(* IEC 61131-3 sources: SortJet_MasterSPS_Aufbau.fbsproj/12_Visu_Uebersicht, 12 files *)

(* ---- VISU_HAND.gvl ---- *)
(* METADATA
{
	"v3Meta": {
		"objectGuid": "6f32179b-dff3-42c9-9870-23893e477a6b"
	}
}
*)
{attribute 'qualified_only'}
NAMESPACE VISU_HAND
VAR_GLOBAL
  st201  : VisuHand_Station_ST;
  st202  : VisuHand_Station_ST;
  st203  : VisuHand_Station_ST;
  st204  : VisuHand_Station_ST;
  st205  : VisuHand_Station_ST;
  st206  : VisuHand_Station_ST;
  st207  : VisuHand_Station_ST;
  st208  : VisuHand_Station_ST;
  st101  : VisuHand_Station_ST;
  st102  : VisuHand_Station_ST;
  st151  : VisuHand_Station_ST;
  st152  : VisuHand_Station_ST;
  astFW  : ARRAY[301..305] OF VisuHand_Station_ST;

  bAnlageResetTaster : BOOL;          // Visu-Taster Anlagen-Reset (einfacher Druck)
  bAnlageResetAktiv  : BOOL;          // Reset laeuft (min. 1 s angezeigt, solange eine Station noch bReset hat)
  sAnlageReset       : STRING(40) := 'ANLAGE RESET';
  dwAnlageResetFarbe : DWORD := 16#FFD64545;
  sLblReset          : STRING(20) := 'Reset';

  // Beschriftungen der Visu "Handbetrieb" (benannt, damit Visu und GVL nicht unbemerkt auseinanderlaufen)
  sL_Riemen                                : STRING(120) := 'Riemen';
  sL_Riemen_X                              : STRING(120) := 'Riemen X';
  sL_Riemen_Y                              : STRING(120) := 'Riemen Y';
  sL_Zur_Zurueck                           : STRING(120) := '<< Zurück';
  sL_Vor_Vor                               : STRING(120) := 'Vor >>';
  sL_Anschlag                              : STRING(120) := 'Anschlag';
  sL_Ab                                    : STRING(120) := 'Ab';
  sL_Auf                                   : STRING(120) := 'Auf';
  sL_Hubrahmen                             : STRING(120) := 'Hubrahmen';
  sL_Senken                                : STRING(120) := 'Senken';
  sL_Heben                                 : STRING(120) := 'Heben';
  sL_Messachse                             : STRING(120) := 'Messachse';
  sL_Minus_Ab                              : STRING(120) := '- Ab';
  sL_Plus_Auf                              : STRING(120) := '+ Auf';
  sL_Referenz                              : STRING(120) := 'Referenz';
  sL_Geblaese                              : STRING(120) := 'Gebläse';
  sL_Ein_Aus                               : STRING(120) := 'Ein / Aus';
  sL_Drosselkl                             : STRING(120) := 'Drosselkl.';
  sL_Auf_Zu                                : STRING(120) := 'Auf / Zu';
  sL_Kippen                                : STRING(120) := 'Kippen';
  sL_Waagerecht                            : STRING(120) := 'Waagerecht';
  sL_Senkrecht                             : STRING(120) := 'Senkrecht';
  sL_Querfahrt                             : STRING(120) := 'Querfahrt';
  sL_Minus_Minus                           : STRING(120) := '- Minus';
  sL_Plus_Plus                             : STRING(120) := '+ Plus';
  sL_84Grad                                : STRING(120) := '84°';
  sL_90Grad                                : STRING(120) := '90°';
  sL_Schmierung                            : STRING(120) := 'Schmierung';
  sL_Starten                               : STRING(120) := 'Starten';
  sL_Riemen_Hub                            : STRING(120) := 'Riemen Hub';
  sL_Anheben                               : STRING(120) := 'Anheben';
  sL_Abfr_Einl                             : STRING(120) := 'Abfr. Einl.';
  sL_Luft_ein                              : STRING(120) := 'Luft ein';
  sL_Abfr_Ausl                             : STRING(120) := 'Abfr. Ausl.';
  sL_Rolltor                               : STRING(120) := 'Rolltor';
  sL_Runter                                : STRING(120) := 'Runter';
  sL_Hoch                                  : STRING(120) := 'Hoch';
  sL_Linearein                             : STRING(120) := 'Linearein.';
  sL_Zurueck                               : STRING(120) := 'Zurück';
  sL_Vor                                   : STRING(120) := 'Vor';
  sL_Shuttle                               : STRING(120) := 'Shuttle';
  sL_Greifer                               : STRING(120) := 'Greifer';
  sL_Oeffnen                               : STRING(120) := 'Öffnen';
  sL_Schliessen                            : STRING(120) := 'Schließen';
  sL_Entriegel                             : STRING(120) := 'Entriegel.';
  sL_Gegenhalter                           : STRING(120) := 'Gegenhalter';
  sL_Lichtschr                             : STRING(120) := 'Lichtschr.';
  sL_Quittieren                            : STRING(120) := 'Quittieren';
  sL_Oeffnung                              : STRING(120) := 'Öffnung';
  sL_16mm                                  : STRING(120) := '16 mm';
  sL_23mm                                  : STRING(120) := '23 mm';
  sL_29mm                                  : STRING(120) := '29 mm';
  sL_Greiferachse                          : STRING(120) := 'Gr.-Achse';
  sL_Zange                                 : STRING(120) := 'Zange';
  sL_Rueckhalter                           : STRING(120) := 'Rückhalter';
  sL_Drehen                                : STRING(120) := 'Drehen';
  sL_0Grad                                 : STRING(120) := '0°';
  sL_180Grad                               : STRING(120) := '180°';
  sL_270Grad                               : STRING(120) := '270°';
  sL_Arretierung                           : STRING(120) := 'Arretierung';
  sL_Einfahren                             : STRING(120) := 'Einfahren';
  sL_Ausfahren                             : STRING(120) := 'Ausfahren';
  sL_Abschrankung                          : STRING(120) := 'Abschrank.';
  sL_HANDBETRIEB                           : STRING(120) := 'HANDBETRIEB';
  sL_Legende                               : STRING(120) := 'Taster (weiß) = Tippbetrieb solange gedrückt   |   Schalter (blau hinterlegt wenn EIN) = Ein/Aus   |   Gesperrt = grau';
  sL_Titel                                 : STRING(120) := 'SortJet  -  Handbetrieb 201 - 208';
  sL_Titel2                                : STRING(120) := 'SortJet  -  Handbetrieb Speicher';
END_VAR
END_NAMESPACE

(* ---- VISU_UEBERSICHT.gvl ---- *)
(* METADATA
{
	"v3Meta": {
		"objectGuid": "76464f8f-3613-4465-9c50-3e0a0f70c8ba"
	}
}
*)
{attribute 'qualified_only'}
NAMESPACE VISU_UEBERSICHT
VAR_GLOBAL
  // Kopfzeile / Anlagenstatus
  sTitel            : STRING(80) := 'SortJet -  Anlagenübersicht';
  sUntertitel       : STRING(120) := 'Anlegetisch 201/205 > Eckübergabe 204 > Drehstation 207 > Shuttle 101 > Speicher > Shuttle 102 > Fächerwagen';
  stAutomatik       : VisuUeb_Lampe_ST;
  stSK1             : VisuUeb_Lampe_ST;
  stSK2             : VisuUeb_Lampe_ST;
  stSK3             : VisuUeb_Lampe_ST;
  stSK4             : VisuUeb_Lampe_ST;
  astTuer               : ARRAY[1..cMAX_TUEREN] OF VisuUeb_Lampe_ST;      // je Tuer eine Anzeige
  abTuerVorhanden       : ARRAY[1..cMAX_TUEREN] OF BOOL;
  astDurchgang          : ARRAY[1..cMAX_DURCHGAENGE] OF VisuUeb_Lampe_ST;
  abDurchgangVorhanden  : ARRAY[1..cMAX_DURCHGAENGE] OF BOOL;
  sLblTueren            : STRING(20) := 'TÜREN';
  sLblDurchgaenge       : STRING(20) := 'DURCHGÄNGE';
  stDruckluft       : VisuUeb_Lampe_ST;
  stSchaltschrank   : VisuUeb_Lampe_ST;
  stEtherCAT        : VisuUeb_Lampe_ST;
  stInit            : VisuUeb_Lampe_ST;
  stMMI             : VisuUeb_Lampe_ST;
  stBetriebsstop    : VisuUeb_Lampe_ST;
  stInbetriebnahme  : VisuUeb_Lampe_ST;
  sStoerungen       : STRING(80);
  dwStoerungenFarbe : DWORD := 16#FF2EAD5B;

  // Stationen
  st501             : VisuUeb_Station_ST;
  st201             : VisuUeb_Station_ST;
  st202             : VisuUeb_Station_ST;
  st203             : VisuUeb_Station_ST;
  st204             : VisuUeb_Station_ST;
  st205             : VisuUeb_Station_ST;
  st206             : VisuUeb_Station_ST;
  st207             : VisuUeb_Station_ST;
  st208             : VisuUeb_Station_ST;
  st101             : VisuUeb_Station_ST;
  st102             : VisuUeb_Station_ST;
  st151             : VisuUeb_Station_ST;
  st152             : VisuUeb_Station_ST;
  st301             : VisuUeb_Station_ST;
  st302             : VisuUeb_Station_ST;
  st303             : VisuUeb_Station_ST;
  st304             : VisuUeb_Station_ST;
  st305             : VisuUeb_Station_ST;

  // Achsen (Querfahrt)
  stAchse101        : VisuUeb_Achse_ST;
  stAchse102        : VisuUeb_Achse_ST;
  stAchse151        : VisuUeb_Achse_ST;
  stAchse152        : VisuUeb_Achse_ST;

  // feste Beschriftungen (Visu nutzt ausschließlich Textvariablen)
  sLblSensoren      : STRING(40) := 'E       EV      AV       A';
  sLblSpeicher      : STRING(40) := 'S O R T I E R S P E I C H E R';
  sLblShuttle101    : STRING(40) := 'SHUTTLE 101';
  sLblTS151         : STRING(40) := 'TRANSFERSHUTTLE 151';
  sLblReset         : STRING(40) := 'Skalierung neu lernen';
  sLblLegende       : STRING(120) := 'Grün = Automatik    Orange = Hand    Blau = Reset / Referenz    Rot = Störung    Grau = deaktiviert';
  sLblNotHaltOK     : STRING(40) := 'NOT-HALT OK';
  sLblNotHaltAus    : STRING(40) := 'NOT-HALT AUSGELÖST';
  sLblStatus        : STRING(40) := 'ANLAGENSTATUS';
  sLblQuerfahrt     : STRING(40) := 'QUERFAHRT';
  sLblIst           : STRING(20) := 'Ist';
  sLblZiel          : STRING(20) := 'Ziel';
  sLblSpeed         : STRING(20) := 'v';
  sLblE             : STRING(4)  := 'E';
  sLblEV            : STRING(4)  := 'EV';
  sLblAV            : STRING(4)  := 'AV';
  sLblA             : STRING(4)  := 'A';
  sLblAS            : STRING(4)  := 'AS';
  sLblQuer101       : STRING(60) := 'QUERFAHRT SHUTTLE 101';
  sLblQuer102       : STRING(60) := 'QUERFAHRT SHUTTLE 102';
  sLblWagen101      : STRING(20) := '101';
  sLblWagen102      : STRING(20) := '102';
  sLblZielMarke     : STRING(10) := 'ZIEL';

  // Bedienung
  bSkalierungNeuLernen : BOOL;
END_VAR

VAR_GLOBAL RETAIN
  // Selbstlernende Skalierung der Fahrbahnen (min/max beobachtete Position)
  bSkalierung101Init : BOOL;
  rMin101            : REAL;
  rMax101            : REAL;
  bSkalierung102Init : BOOL;
  rMin102            : REAL;
  rMax102            : REAL;
  bSkalierung151Init : BOOL;
  rMin151            : REAL;
  rMax151            : REAL;
  bSkalierung152Init : BOOL;
  rMin152            : REAL;
  rMax152            : REAL;
END_VAR

VAR_GLOBAL CONSTANT
  cMAX_TUEREN          : WORD := 8;     // Anzahl Tueranzeigen in der Visu
  cMAX_DURCHGAENGE     : WORD := 3;     // Anzahl Durchganganzeigen in der Visu
  cBAHN_LAENGE_PX      : INT  := 266;   // nutzbare Laenge der senkrechten Fahrbahn (muss zur Visu passen)
  cWAGEN_LAENGE_PX     : INT  := 34;    // Hoehe Fahrwagen (muss zur Visu passen)
  cMIN_SPANNE_MM       : REAL := 500;   // minimale Skalierungsspanne

  cFARBE_GRUEN         : DWORD := 16#FF2EAD5B;
  cFARBE_ROT           : DWORD := 16#FFD64545;
  cFARBE_ORANGE        : DWORD := 16#FFF0A202;
  cFARBE_BLAU          : DWORD := 16#FF2F80ED;
  cFARBE_GRAU          : DWORD := 16#FF9AA5B1;
  cFARBE_GRAU_HELL     : DWORD := 16#FFE4E7EB;
  cFARBE_RAHMEN        : DWORD := 16#FFCBD2D9;
  cFARBE_TEXT          : DWORD := 16#FF52606D;
  cFARBE_SENSOR_AN     : DWORD := 16#FFFFC531;
END_VAR
END_NAMESPACE

(* ---- VisuHand_Set.fn.st ---- *)
(* METADATA
{
	"v3Meta": {
		"objectGuid": "443bc09b-b8af-4511-9c3a-ed00ec4cc080"
	}
}
*)
FUNCTION VisuHand_Set : BOOL
VAR_IN_OUT
  stH     : VisuHand_Station_ST;
END_VAR
VAR_INPUT
  wZeile  : WORD;
  sText   : STRING(30);
  dwFarbe : DWORD;
END_VAR
IF wZeile >= 1 AND wZeile <= 10 THEN // Grenzen wie VisuHand_Station_ST.asStatus
  stH.asStatus[wZeile]  := sText;
  stH.adwStatus[wZeile] := dwFarbe;
END_IF
VisuHand_Set := TRUE;
END_FUNCTION

(* ---- VisuHand_Sperre.fn.st ---- *)
(* METADATA
{
	"v3Meta": {
		"objectGuid": "d31da620-9df0-4563-ab06-3d7039f98cd3"
	}
}
*)
FUNCTION VisuHand_Sperre : BOOL
VAR_IN_OUT
  stBP : StationBasisParameter_ST;
  stH  : VisuHand_Station_ST;
END_VAR
VAR_INPUT
  bFaecherwagen : BOOL; // FW-Handfunktionen sind im FB nicht an die Betriebsart gebunden -> hier zusaetzlich bei Automatik sperren
END_VAR
VAR
  bDeaktiviert : BOOL;
END_VAR
IF __ISVALIDREF(stBP.stMKs) THEN
  bDeaktiviert := stBP.stMKs.bDeaktivieren;
END_IF

IF bDeaktiviert THEN
  stH.bGesperrt := TRUE;  stH.sSperrgrund := 'Gesperrt: Station deaktiviert';
ELSIF stBP.bAutomatik THEN
  stH.bGesperrt := TRUE;  stH.sSperrgrund := 'Gesperrt: Automatik aktiv';
ELSIF stBP.bReset THEN
  stH.bGesperrt := TRUE;  stH.sSperrgrund := 'Gesperrt: Reset läuft';
ELSIF stBP.bReferenz THEN
  stH.bGesperrt := TRUE;  stH.sSperrgrund := 'Gesperrt: Referenzfahrt läuft';
ELSIF stBP.bCheck THEN
  stH.bGesperrt := TRUE;  stH.sSperrgrund := 'Gesperrt: Systemcheck läuft';
ELSIF bFaecherwagen AND (stBP.bEintransport[cWAND_1] OR stBP.bAustransport[cWAND_1]) THEN
  stH.bGesperrt := TRUE;  stH.sSperrgrund := 'Gesperrt: Ein-/Ausschleusen aktiv';
ELSE
  stH.bGesperrt := FALSE;
  stH.sSperrgrund := SEL(stBP.stFreigabe.bAlles, 'Hand frei - keine Sicherheitsfreigabe', 'Handbetrieb freigegeben');
END_IF

IF stH.bGesperrt THEN
  stH.dwSperrFarbe := VISU_UEBERSICHT.cFARBE_GRAU;
ELSIF NOT stBP.stFreigabe.bAlles THEN
  stH.dwSperrFarbe := VISU_UEBERSICHT.cFARBE_ORANGE;
ELSE
  stH.dwSperrFarbe := VISU_UEBERSICHT.cFARBE_GRUEN;
END_IF
VisuHand_Sperre := stH.bGesperrt;
END_FUNCTION

(* ---- VisuUeb_Achse.fn.st ---- *)
(* METADATA
{
	"v3Meta": {
		"objectGuid": "3979691c-e077-4914-8fb4-604417bd71fb"
	}
}
*)
FUNCTION VisuUeb_Achse : BOOL
VAR_IN_OUT
  stAchse   : VisuUeb_Achse_ST;
  bInit     : BOOL;  // Skalierung initialisiert (RETAIN)
  rMin      : REAL;  // gelerntes Minimum (RETAIN)
  rMax      : REAL;  // gelerntes Maximum (RETAIN)
END_VAR
VAR_INPUT
  rIst         : REAL;
  rZiel        : REAL;
  rSpeed       : REAL;
  bPositionierung : BOOL;
  bReferenziert   : BOOL;
  bFehler         : BOOL;
  bMinEnd         : BOOL;
  bMaxEnd         : BOOL;
  bNeuLernen      : BOOL;
  bBlink          : BOOL;
  rSkalaMin       : REAL;  // gemeinsamer Darstellungsbereich mehrerer Achsen (Max <= Min: eigener Bereich)
  rSkalaMax       : REAL;
END_VAR
VAR
  rSpanne : REAL;
  rFaktor : REAL;
  iWeg    : INT;
  rDarstMin : REAL;
END_VAR
// Skalierung lernen (nur mit gueltiger Referenz)
IF bNeuLernen THEN
  bInit := FALSE;
END_IF
IF bReferenziert THEN
  IF NOT bInit THEN
    rMin  := rIst;
    rMax  := rIst;
    bInit := TRUE;
  END_IF
  rMin := MIN(rMin, rIst);
  rMax := MAX(rMax, rIst);
  IF bPositionierung THEN
    rMin := MIN(rMin, rZiel);
    rMax := MAX(rMax, rZiel);
  END_IF
END_IF

IF rSkalaMax > rSkalaMin THEN
  rDarstMin := rSkalaMin;
  rSpanne   := MAX(rSkalaMax - rSkalaMin, VISU_UEBERSICHT.cMIN_SPANNE_MM);
ELSE
  rDarstMin := rMin;
  rSpanne   := MAX(rMax - rMin, VISU_UEBERSICHT.cMIN_SPANNE_MM);
END_IF
iWeg    := VISU_UEBERSICHT.cBAHN_LAENGE_PX - VISU_UEBERSICHT.cWAGEN_LAENGE_PX;

rFaktor := LIMIT(0.0, (rIst - rDarstMin) / rSpanne, 1.0);
stAchse.iPixel := REAL_TO_INT(rFaktor * INT_TO_REAL(iWeg));
rFaktor := LIMIT(0.0, (rZiel - rDarstMin) / rSpanne, 1.0);
stAchse.iZielPixel := REAL_TO_INT(rFaktor * INT_TO_REAL(iWeg));

stAchse.rIstPos         := rIst;
stAchse.rZielPos        := rZiel;
stAchse.rSpeed          := rSpeed;
stAchse.bPositionierung := bPositionierung;
stAchse.bReferenziert   := bReferenziert;
stAchse.sIstPos         := VisuUeb_MmText(sPrefix := 'Ist  ', rWert := rIst);
stAchse.sZielPos        := SEL(bPositionierung, 'Ziel  -', VisuUeb_MmText(sPrefix := 'Ziel  ', rWert := rZiel));
stAchse.sSpeed          := VisuUeb_MmText(sPrefix := 'v  ', rWert := rSpeed, sEinheit := ' mm/s');
stAchse.sBereich        := CONCAT(CONCAT(VisuUeb_MmText(sPrefix := 'Bereich ', rWert := rMin), ' ... '), VisuUeb_MmText(sPrefix := '', rWert := rMax));

IF bFehler THEN
  stAchse.dwKoerperFarbe := SEL(bBlink, 16#FF8C2F2F, VISU_UEBERSICHT.cFARBE_ROT);
ELSIF NOT bReferenziert THEN
  stAchse.dwKoerperFarbe := VISU_UEBERSICHT.cFARBE_ORANGE;
ELSIF bPositionierung THEN
  stAchse.dwKoerperFarbe := 16#FF1C64CC;
ELSE
  stAchse.dwKoerperFarbe := VISU_UEBERSICHT.cFARBE_BLAU;
END_IF
stAchse.dwMinEndFarbe := SEL(bMinEnd, VISU_UEBERSICHT.cFARBE_GRAU_HELL, VISU_UEBERSICHT.cFARBE_ROT);
stAchse.dwMaxEndFarbe := SEL(bMaxEnd, VISU_UEBERSICHT.cFARBE_GRAU_HELL, VISU_UEBERSICHT.cFARBE_ROT);
VisuUeb_Achse := bInit;
END_FUNCTION

(* ---- VisuUeb_Lampe.fn.st ---- *)
(* METADATA
{
	"v3Meta": {
		"objectGuid": "b7aa09e8-5cde-43cf-b09b-dc0ab15a15f2"
	}
}
*)
FUNCTION VisuUeb_Lampe : BOOL
VAR_IN_OUT
  stLampe   : VisuUeb_Lampe_ST;
END_VAR
VAR_INPUT
  sText     : STRING(40);
  bOK       : BOOL;   // TRUE = gruen
  bWarnung  : BOOL := FALSE; // bei NOT bOK: TRUE = orange, FALSE = rot
  bNeutral  : BOOL := FALSE; // TRUE = grau (inaktiv, keine Bewertung)
END_VAR
stLampe.sText := sText;
IF bNeutral THEN
  stLampe.dwFarbe := VISU_UEBERSICHT.cFARBE_GRAU;
ELSIF bOK THEN
  stLampe.dwFarbe := VISU_UEBERSICHT.cFARBE_GRUEN;
ELSIF bWarnung THEN
  stLampe.dwFarbe := VISU_UEBERSICHT.cFARBE_ORANGE;
ELSE
  stLampe.dwFarbe := VISU_UEBERSICHT.cFARBE_ROT;
END_IF
VisuUeb_Lampe := bOK;
END_FUNCTION

(* ---- VisuUeb_MmText.fn.st ---- *)
(* METADATA
{
	"v3Meta": {
		"objectGuid": "478effab-2bb6-4cba-a63b-7b7e6c506f75"
	}
}
*)
FUNCTION VisuUeb_MmText : STRING(40)
VAR_INPUT
  sPrefix : STRING(20);
  rWert   : REAL;
  sEinheit: STRING(10) := ' mm';
END_VAR
VisuUeb_MmText := CONCAT(CONCAT(sPrefix, DINT_TO_STRING(REAL_TO_DINT(rWert))), sEinheit);
END_FUNCTION

(* ---- VisuUeb_Sensor.fn.st ---- *)
(* METADATA
{
	"v3Meta": {
		"objectGuid": "2f1f2564-8eff-43f7-8c8f-4a939be6a082"
	}
}
*)
FUNCTION VisuUeb_Sensor : DWORD
VAR_INPUT
  bBelegt    : BOOL;
  bVorhanden : BOOL := TRUE;
END_VAR
IF NOT bVorhanden THEN
  VisuUeb_Sensor := 16#00FFFFFF; // transparent
ELSIF bBelegt THEN
  VisuUeb_Sensor := VISU_UEBERSICHT.cFARBE_SENSOR_AN;
ELSE
  VisuUeb_Sensor := VISU_UEBERSICHT.cFARBE_GRAU_HELL;
END_IF
END_FUNCTION

(* ---- VisuUeb_Station.fn.st ---- *)
(* METADATA
{
	"v3Meta": {
		"objectGuid": "2a69d02d-507f-4a31-bfce-f3b7167a1195"
	}
}
*)
FUNCTION VisuUeb_Station : BOOL
VAR_IN_OUT
  stBP    : StationBasisParameter_ST;
  stKarte : VisuUeb_Station_ST;
END_VAR
VAR_INPUT
  sTitel  : STRING(40);
  bBlink  : BOOL;
  bGlasZusatz : BOOL := FALSE; // zusaetzliche Glaserkennung (z.B. Sensoren)
  bReferenzRelevant : BOOL := TRUE; // FALSE: Station hat keine referenzierbaren Achsen (z.B. Faecherwagen)
END_VAR
VAR
  bDeaktiviert : BOOL;
END_VAR
stKarte.sTitel := sTitel;
IF __ISVALIDREF(stBP.stMKs) THEN
  bDeaktiviert := stBP.stMKs.bDeaktivieren;
END_IF
stKarte.bDeaktiviert := bDeaktiviert;

// Referenzstatus (BasisStationsParameter.bIstReferenziert)
stKarte.bReferenzAnzeigen := bReferenzRelevant AND NOT bDeaktiviert;
IF stBP.bIstReferenziert THEN
  stKarte.sReferenz := 'REFERENZIERT';      stKarte.dwReferenzFarbe := VISU_UEBERSICHT.cFARBE_GRUEN;
ELSIF stBP.bReferenz THEN
  stKarte.sReferenz := 'REFERENZIERT ...';  stKarte.dwReferenzFarbe := SEL(bBlink, VISU_UEBERSICHT.cFARBE_GRAU, VISU_UEBERSICHT.cFARBE_BLAU);
ELSE
  stKarte.sReferenz := 'NICHT REFERENZIERT'; stKarte.dwReferenzFarbe := VISU_UEBERSICHT.cFARBE_ORANGE;
END_IF

// Zustand
IF bDeaktiviert THEN
  stKarte.sZustand := 'DEAKTIVIERT';         stKarte.dwZustandFarbe := VISU_UEBERSICHT.cFARBE_GRAU;
ELSIF stBP.bFehler THEN
  stKarte.sZustand := 'STÖRUNG';             stKarte.dwZustandFarbe := VISU_UEBERSICHT.cFARBE_ROT;
ELSIF stBP.bReset THEN
  stKarte.sZustand := 'RESET';               stKarte.dwZustandFarbe := VISU_UEBERSICHT.cFARBE_BLAU;
ELSIF stBP.bReferenz THEN
  stKarte.sZustand := 'REFERENZFAHRT';       stKarte.dwZustandFarbe := VISU_UEBERSICHT.cFARBE_BLAU;
ELSIF stBP.bCheck THEN
  stKarte.sZustand := 'SYSTEMCHECK';         stKarte.dwZustandFarbe := VISU_UEBERSICHT.cFARBE_BLAU;
ELSIF stBP.bAutomatik THEN
  stKarte.sZustand := 'AUTOMATIK';           stKarte.dwZustandFarbe := VISU_UEBERSICHT.cFARBE_GRUEN;
ELSE
  stKarte.sZustand := 'HAND';                stKarte.dwZustandFarbe := VISU_UEBERSICHT.cFARBE_ORANGE;
END_IF

// Rahmen: Stoerung blinkt rot, aktiver Auftrag blau
IF stBP.bFehler AND NOT bDeaktiviert THEN
  stKarte.dwRahmenFarbe := SEL(bBlink, VISU_UEBERSICHT.cFARBE_RAHMEN, VISU_UEBERSICHT.cFARBE_ROT);
ELSIF stBP.bAuftragAktiv THEN
  stKarte.dwRahmenFarbe := VISU_UEBERSICHT.cFARBE_BLAU;
ELSE
  stKarte.dwRahmenFarbe := VISU_UEBERSICHT.cFARBE_RAHMEN;
END_IF

// Aktive Funktion
IF bDeaktiviert THEN
  stKarte.sFunktion := '-';
ELSIF stBP.bFehler THEN
  stKarte.sFunktion := CONCAT('Fehlernummer ', WORD_TO_STRING(stBP.wFehlerNummer));
ELSIF stBP.bAnlegen THEN                      stKarte.sFunktion := 'Anlegen';
ELSIF stBP.bAbnehmen THEN                     stKarte.sFunktion := 'Abnehmen';
ELSIF stBP.bEintransport[cWAND_1] THEN        stKarte.sFunktion := 'Eintransport';
ELSIF stBP.bAustransport[cWAND_1] THEN        stKarte.sFunktion := 'Austransport';
ELSIF stBP.bDurchtransport[cWAND_1] THEN      stKarte.sFunktion := 'Durchtransport';
ELSIF stBP.bVortransport[cWAND_1] THEN        stKarte.sFunktion := 'Vortransport';
ELSIF stBP.bTransportkopplung[cWAND_1] THEN   stKarte.sFunktion := 'Transportkopplung';
ELSIF stBP.bMesskopplung[cWAND_1] THEN        stKarte.sFunktion := 'Messkopplung';
ELSIF stBP.bGlaslaengenmessung THEN           stKarte.sFunktion := 'Glaslängenmessung';
ELSIF stBP.bGlashoehenmessung THEN            stKarte.sFunktion := 'Glashöhenmessung';
ELSIF stBP.bVorabpositionieren THEN           stKarte.sFunktion := 'Vorabpositionierung';
ELSIF stBP.bAuftragAktiv THEN                 stKarte.sFunktion := 'Auftrag aktiv';
ELSIF stBP.stFreigabe.bAlles THEN                     stKarte.sFunktion := 'Bereit';
ELSE                                          stKarte.sFunktion := 'Keine Freigabe';
END_IF

stKarte.bGlas := stBP.bStationBelegt[cWAND_1] OR bGlasZusatz;
VisuUeb_Station := stBP.bFehler AND NOT bDeaktiviert;
END_FUNCTION

(* ---- VisuHand_Reset_FB.fb.st ---- *)
(* METADATA
{
	"v3Meta": {
		"objectGuid": "8e79010e-8dea-435f-8304-0b4307ea198e"
	}
}
*)
FUNCTION_BLOCK VisuHand_Reset_FB
// Stations-Reset aus der Visu:
//   - setzt BasisStationsParameter.bReset (die Station fuehrt ihre eigene Reset-Aktion aus und setzt bReset selbst zurueck)
//   - nur ausserhalb der Automatik, nicht wenn die Station deaktiviert ist oder bereits ein Reset laeuft
VAR_IN_OUT
  stBP : StationBasisParameter_ST;
  stH  : VisuHand_Station_ST;
END_VAR
VAR
  rtlTaster    : R_TRIG;
  bDeaktiviert : BOOL;
END_VAR
bDeaktiviert := FALSE;
IF __ISVALIDREF(stBP.stMKs) THEN
  bDeaktiviert := stBP.stMKs.bDeaktivieren;
END_IF

stH.bResetGesperrt := bDeaktiviert OR stBP.bAutomatik OR stBP.bReset OR stBP.bReferenz OR stBP.bCheck;

rtlTaster(CLK := stH.bResetTaster);
IF rtlTaster.Q AND NOT stH.bResetGesperrt THEN
  stBP.bReset := TRUE;
END_IF
END_FUNCTION_BLOCK

(* ---- VisuHand_PRG.prg.st ---- *)
(* METADATA
{
	"v3Meta": {
		"objectGuid": "a4fab899-80a6-4d8b-aad2-f00973a33795"
	}
}
*)
PROGRAM VisuHand_PRG
VAR
  b    : BOOL;
  i    : WORD;
  dwG, dwO, dwR, dwGR, dwB : DWORD;
  sKipp : STRING(30);
  dwKipp : DWORD;
  pBP  : POINTER TO StationBasisParameter_ST;
  pH   : POINTER TO VisuHand_Station_ST;
  pGr  : POINTER TO Shuttle_Greifer_FB_V01_00_00; // Greifer Wand 1 des Shuttles (Zeilen 7 - 10)

  // Reset
  afbResetSt       : ARRAY[201..208] OF VisuHand_Reset_FB;
  afbResetSh       : ARRAY[101..102] OF VisuHand_Reset_FB;
  afbResetTS       : ARRAY[151..152] OF VisuHand_Reset_FB;
  afbResetFW       : ARRAY[301..305] OF VisuHand_Reset_FB;
  rtlAnlageReset   : R_TRIG;  // Anlagen-Reset auf Flanke
  tofAnlageReset   : TOF;     // Mindestanzeige "Reset aktiv"
  bResetLaeuft     : BOOL;

  // Rolltor-Schalter (Toggle) gegenseitig ausschliessen
  artlRolltorHoch, artlRolltorRunter : ARRAY[301..305] OF R_TRIG;
END_VAR
// *************************************************************************************************
// DATENAUFBEREITUNG FUER DIE VISUS "Handbetrieb" (201 - 208) UND "Handbetrieb_Speicher"
// (Shuttle 101/102, Transfershuttle 151/152, Faecherwagen 301 - 305)
// - Taster schreiben direkt auf die vorhandenen VISU_VARS-Bits
// - hier nur: Sperre je Station + Rueckmeldetexte/-farben
// *************************************************************************************************
dwG  := VISU_UEBERSICHT.cFARBE_GRUEN;
dwO  := VISU_UEBERSICHT.cFARBE_ORANGE;
dwR  := VISU_UEBERSICHT.cFARBE_ROT;
dwGR := VISU_UEBERSICHT.cFARBE_GRAU;
dwB  := VISU_UEBERSICHT.cFARBE_BLAU;

// -------------------------------------------------------------------------------------------
// RESET
// - Anlage: wie "Stopp" vom MMI (alle Automatikkreise stoppen + Reset aller Stationen)
// - Station: BasisStationsParameter.bReset (nur ausserhalb der Automatik)
// -------------------------------------------------------------------------------------------
rtlAnlageReset(CLK := VISU_HAND.bAnlageResetTaster);
IF rtlAnlageReset.Q THEN
  MMI_Vars.tMmi2SpsInfo.wAutomatikStopArea   := Stations_Konfig.cSTOPP_ALLE_AUTOMATIKKREIS;
  MMI_Vars.M_SB0_MMI_SortierungAutomatik_Stop := TRUE;
END_IF

bResetLaeuft := FALSE;
FOR i := 201 TO 208 DO
  CASE i OF
    201: pH := ADR(VISU_HAND.st201);
    202: pH := ADR(VISU_HAND.st202);
    203: pH := ADR(VISU_HAND.st203);
    204: pH := ADR(VISU_HAND.st204);
    205: pH := ADR(VISU_HAND.st205);
    206: pH := ADR(VISU_HAND.st206);
    207: pH := ADR(VISU_HAND.st207);
    208: pH := ADR(VISU_HAND.st208);
  END_CASE
  afbResetSt[i](stBP := StationBasisParameter.starrStationBasisParameter[i], stH := pH^);
  bResetLaeuft := bResetLaeuft OR StationBasisParameter.starrStationBasisParameter[i].bReset;
END_FOR
afbResetSh[101](stBP := StationBasisParameter.starrShuttleBasisParameter[101], stH := VISU_HAND.st101);
afbResetSh[102](stBP := StationBasisParameter.starrShuttleBasisParameter[102], stH := VISU_HAND.st102);
afbResetTS[151](stBP := StationBasisParameter.starrTransfershuttleBasisParameter[151], stH := VISU_HAND.st151);
afbResetTS[152](stBP := StationBasisParameter.starrTransfershuttleBasisParameter[152], stH := VISU_HAND.st152);
FOR i := 101 TO 102 DO
  bResetLaeuft := bResetLaeuft OR StationBasisParameter.starrShuttleBasisParameter[i].bReset;
END_FOR
FOR i := 151 TO 152 DO
  bResetLaeuft := bResetLaeuft OR StationBasisParameter.starrTransfershuttleBasisParameter[i].bReset;
END_FOR
FOR i := 301 TO 305 DO
  afbResetFW[i](stBP := StationBasisParameter.starrFaecherwagenBasisParameter[i], stH := VISU_HAND.astFW[i]);
  bResetLaeuft := bResetLaeuft OR StationBasisParameter.starrFaecherwagenBasisParameter[i].bReset;
END_FOR

// Reset aktiv: min. 1 s nach Druck bzw. solange irgendeine Station ihren Reset noch nicht abgeschlossen hat
tofAnlageReset(IN := rtlAnlageReset.Q, PT := T#1S);
VISU_HAND.bAnlageResetAktiv := tofAnlageReset.Q OR bResetLaeuft;
IF VISU_HAND.bAnlageResetAktiv THEN
  VISU_HAND.sAnlageReset       := 'RESET AKTIV ...';
  VISU_HAND.dwAnlageResetFarbe := dwO;
ELSE
  VISU_HAND.sAnlageReset       := 'ANLAGE RESET';
  VISU_HAND.dwAnlageResetFarbe := dwR;
END_IF

// -------------------------------------------------------------------------------------------
// [201] - [208] STATIONEN: Sperre, Funktionszeilen laut MK-Stationsaufbau, Rueckmeldungen
// -------------------------------------------------------------------------------------------
FOR i := 201 TO 208 DO
  CASE i OF
    201: pH := ADR(VISU_HAND.st201);
    202: pH := ADR(VISU_HAND.st202);
    203: pH := ADR(VISU_HAND.st203);
    204: pH := ADR(VISU_HAND.st204);
    205: pH := ADR(VISU_HAND.st205);
    206: pH := ADR(VISU_HAND.st206);
    207: pH := ADR(VISU_HAND.st207);
    208: pH := ADR(VISU_HAND.st208);
  END_CASE
  pBP := ADR(StationBasisParameter.starrStationBasisParameter[i]);
  b := VisuHand_Sperre(stBP := pBP^, stH := pH^, bFaecherwagen := FALSE);

  // Funktionszeilen
  IF __ISVALIDREF(pBP^.stMKs) THEN
    pH^.abZeileVorhanden[1] := pBP^.stMKs.stStationsAufbau.bGlastransport[cWAND_1];
    CASE i OF
      201, 205:
        pH^.abZeileVorhanden[2] := pBP^.stMKs.stStationsAufbau.bAnschlag;
        pH^.abZeileVorhanden[3] := pBP^.stMKs.stStationsAufbau.bHubrahmen;
        pH^.abZeileVorhanden[4] := pBP^.stMKs.stStationsAufbau.bMessachse;
        pH^.abZeileVorhanden[5] := pBP^.stMKs.stStationsAufbau.bGeblase[cWAND_1];
        pH^.abZeileVorhanden[6] := pBP^.stMKs.stStationsAufbau.bGeblase[cWAND_1];
      204:
        pH^.abZeileVorhanden[2] := pBP^.stMKs.stStationsAufbau.bGlastransport[cWAND_1];
        pH^.abZeileVorhanden[3] := pBP^.stMKs.stStationsAufbau.bHubrahmen;
      206:
        pH^.abZeileVorhanden[2] := pBP^.stMKs.stStationsAufbau.bKippen[cWAND_1];
      207:
        pH^.abZeileVorhanden[2] := pBP^.stMKs.stStationsAufbau.bDrehen;
        pH^.abZeileVorhanden[3] := pBP^.stMKs.stStationsAufbau.bDrehen;
        pH^.abZeileVorhanden[4] := pBP^.stMKs.stStationsAufbau.bDrehen;
        pH^.abZeileVorhanden[5] := pBP^.stMKs.stStationsAufbau.bKippen[cWAND_1];
        pH^.abZeileVorhanden[6] := pBP^.stMKs.stStationsAufbau.bGeblase[cWAND_1];
      208:
        pH^.abZeileVorhanden[2] := pBP^.stMKs.stStationsAufbau.bMessachse;
        pH^.abZeileVorhanden[3] := pBP^.stMKs.stStationsAufbau.bDurchlaufSperreZumNachfolger;
    END_CASE
  END_IF

  // 1 Riemen: Glas auf der Station
  b := VisuHand_Set(stH := pH^, wZeile := 1,
                     sText   := SEL(abgStationsstatusVisu[i].bSensorEinlauf[1] OR abgStationsstatusVisu[i].bSensorAuslauf[1], 'frei', 'Glas'),
                     dwFarbe := SEL(abgStationsstatusVisu[i].bSensorEinlauf[1] OR abgStationsstatusVisu[i].bSensorAuslauf[1], dwGR, dwB));

  CASE i OF
    201, 205:
      // 1 Riemen (laeuft nur bei ausgefahrenem Hubrahmen)
      IF NOT abgStationsstatusVisu[i].bHubpaletteSensorAusgefahren THEN
        b := VisuHand_Set(stH := pH^, wZeile := 1, sText := 'Hubr. unten', dwFarbe := dwO);
      END_IF
      // 2 Anschlag
      IF abgStationsstatusVisu[i].bAnschlagFehler THEN                   b := VisuHand_Set(stH := pH^, wZeile := 2, sText := 'Fehler', dwFarbe := dwR);
      ELSIF abgStationsstatusVisu[i].bAnschlagSensorAusgefahren THEN     b := VisuHand_Set(stH := pH^, wZeile := 2, sText := 'oben',   dwFarbe := dwG);
      ELSIF abgStationsstatusVisu[i].bAnschlagSensorEingefahren THEN     b := VisuHand_Set(stH := pH^, wZeile := 2, sText := 'unten',  dwFarbe := dwG);
      ELSE                                                               b := VisuHand_Set(stH := pH^, wZeile := 2, sText := '?',      dwFarbe := dwO);
      END_IF
      // 3 Hubrahmen
      IF abgStationsstatusVisu[i].bHubpaletteFehler THEN                 b := VisuHand_Set(stH := pH^, wZeile := 3, sText := 'Fehler', dwFarbe := dwR);
      ELSIF abgStationsstatusVisu[i].bHubpaletteSensorAusgefahren THEN   b := VisuHand_Set(stH := pH^, wZeile := 3, sText := 'oben',   dwFarbe := dwG);
      ELSIF abgStationsstatusVisu[i].bHubpaletteSensorEingefahren THEN   b := VisuHand_Set(stH := pH^, wZeile := 3, sText := 'unten',  dwFarbe := dwG);
      ELSE                                                               b := VisuHand_Set(stH := pH^, wZeile := 3, sText := '?',      dwFarbe := dwO);
      END_IF
      // 4 Messachse
      b := VisuHand_Set(stH := pH^, wZeile := 4,
                         sText   := VisuUeb_MmText(sPrefix := '', rWert := abgStationsstatusVisu[i].rMessachseIstPos, sEinheit := ' mm'),
                         dwFarbe := SEL(abgStationsstatusVisu[i].bMessachseFehler, SEL(pBP^.bIstReferenziert, dwO, dwG), dwR));
      // 5 Geblaese
      b := VisuHand_Set(stH := pH^, wZeile := 5, sText := SEL(abgStationsstatusVisu[i].bGeblaeseLaeuft[1], 'aus', 'EIN'), dwFarbe := SEL(abgStationsstatusVisu[i].bGeblaeseLaeuft[1], dwGR, dwB));
      // 6 Drosselklappe (Ausgang, keine Endlagenabfrage)
      b := VisuHand_Set(stH := pH^, wZeile := 6, sText := SEL(abgStationsstatusVisu[i].bDrosselklappeOffen[1], 'zu', 'auf'), dwFarbe := SEL(abgStationsstatusVisu[i].bDrosselklappeOffen[1], dwGR, dwB));

    204:
      // 2 Riemen Y: Sensoren nur fuer die X-Achse in der Visu-Schnittstelle
      b := VisuHand_Set(stH := pH^, wZeile := 2, sText := '', dwFarbe := dwGR);
      // 3 Hubrahmen (oben = Riemen X arbeitet)
      IF abgStationsstatusVisu[i].bHubpaletteFehler THEN                 b := VisuHand_Set(stH := pH^, wZeile := 3, sText := 'Fehler', dwFarbe := dwR);
      ELSIF abgStationsstatusVisu[i].bHubpaletteSensorAusgefahren THEN   b := VisuHand_Set(stH := pH^, wZeile := 3, sText := 'oben',   dwFarbe := dwG);
      ELSIF abgStationsstatusVisu[i].bHubpaletteSensorEingefahren THEN   b := VisuHand_Set(stH := pH^, wZeile := 3, sText := 'unten',  dwFarbe := dwG);
      ELSE                                                               b := VisuHand_Set(stH := pH^, wZeile := 3, sText := '?',      dwFarbe := dwO);
      END_IF

    206:
      // 2 Kippen
      CASE abgStationsstatusVisu[i].epKippStatus OF
        Kippen_EN.eKippen_Position_0Grad:    sKipp := 'waagerecht'; dwKipp := dwG;
        Kippen_EN.eKippen_Position_90Grad:   sKipp := 'senkrecht';  dwKipp := dwG;
        Kippen_EN.eKippen_Position_84Grad:   sKipp := '84°';        dwKipp := dwG;
        Kippen_EN.eKippen_Position_88_5Grad: sKipp := '88,5°';      dwKipp := dwG;
        Kippen_EN.eKippen_Position_96Grad:   sKipp := '96°';        dwKipp := dwG;
        Kippen_EN.eKippen_Fehler:            sKipp := 'Fehler';     dwKipp := dwR;
        ELSE                                   sKipp := 'Zwischen';   dwKipp := dwO;
      END_CASE
      IF abgStationsstatusVisu[i].bKippenFehler THEN dwKipp := dwR; ELSIF NOT abgStationsstatusVisu[i].bKippenAntriebReferenziert THEN dwKipp := dwO; END_IF
      b := VisuHand_Set(stH := pH^, wZeile := 2, sText := sKipp, dwFarbe := dwKipp);

    207:
      // 2 Drehen: Position
      CASE abgStationsstatusVisu[i].epDrehIstPosition OF
        Drehen_EN.eDrehPosition0Grad:   sKipp := '0°';   dwKipp := dwG;
        Drehen_EN.eDrehPosition90Grad:  sKipp := '90°';  dwKipp := dwG;
        Drehen_EN.eDrehPosition180Grad: sKipp := '180°'; dwKipp := dwG;
        Drehen_EN.eDrehPosition270Grad: sKipp := '270°'; dwKipp := dwG;
        ELSE                              sKipp := 'Zwischen'; dwKipp := dwO;
      END_CASE
      IF abgStationsstatusVisu[i].bDrehenFehler THEN sKipp := 'Fehler'; dwKipp := dwR; END_IF
      b := VisuHand_Set(stH := pH^, wZeile := 2, sText := sKipp, dwFarbe := dwKipp);
      // 3 Drehen: Referenz
      b := VisuHand_Set(stH := pH^, wZeile := 3,
                         sText   := SEL(abgStationsstatusVisu[i].bDrehenAntriebReferenziert, 'nicht ref.', 'referenz.'),
                         dwFarbe := SEL(abgStationsstatusVisu[i].bDrehenAntriebReferenziert, dwO, dwG));
      // 4 Arretierung
      IF abgStationsstatusVisu[i].bDrehenArretierungAusgefahren THEN
        b := VisuHand_Set(stH := pH^, wZeile := 4, sText := 'ausgefahren', dwFarbe := dwG);
      ELSIF abgStationsstatusVisu[i].bDrehenArretierungEingefahren THEN
        b := VisuHand_Set(stH := pH^, wZeile := 4, sText := 'eingefahren', dwFarbe := dwG);
      ELSE
        b := VisuHand_Set(stH := pH^, wZeile := 4, sText := '?', dwFarbe := dwO);
      END_IF
      // 5 Kippen
      CASE abgStationsstatusVisu[i].epKippStatus OF
        Kippen_EN.eKippen_Position_84Grad: sKipp := '84°';    dwKipp := dwG;
        Kippen_EN.eKippen_Position_90Grad: sKipp := '90°';    dwKipp := dwG;
        Kippen_EN.eKippen_Fehler:          sKipp := 'Fehler'; dwKipp := dwR;
        ELSE                                 sKipp := 'Zwischen'; dwKipp := dwO;
      END_CASE
      IF abgStationsstatusVisu[i].bKippenFehler THEN sKipp := 'Fehler'; dwKipp := dwR; END_IF
      b := VisuHand_Set(stH := pH^, wZeile := 5, sText := sKipp, dwFarbe := dwKipp);
      // 6 Geblaese
      b := VisuHand_Set(stH := pH^, wZeile := 6, sText := SEL(abgStationsstatusVisu[i].bGeblaeseLaeuft[1], 'aus', 'EIN'), dwFarbe := SEL(abgStationsstatusVisu[i].bGeblaeseLaeuft[1], dwGR, dwB));

    208:
      // 2 Messachse
      b := VisuHand_Set(stH := pH^, wZeile := 2,
                         sText   := VisuUeb_MmText(sPrefix := '', rWert := abgStationsstatusVisu[i].rMessachseIstPos, sEinheit := ' mm'),
                         dwFarbe := SEL(abgStationsstatusVisu[i].bMessachseFehler, SEL(pBP^.bIstReferenziert, dwO, dwG), dwR));
      // 3 Bewegliche Abschrankung
      IF abgStationsstatusVisu[i].bAbschrankungFehler THEN             b := VisuHand_Set(stH := pH^, wZeile := 3, sText := 'Fehler', dwFarbe := dwR);
      ELSIF abgStationsstatusVisu[i].bAbschrankungGeschlossen THEN     b := VisuHand_Set(stH := pH^, wZeile := 3, sText := 'zu',     dwFarbe := dwG);
      ELSIF abgStationsstatusVisu[i].bAbschrankungOffen THEN           b := VisuHand_Set(stH := pH^, wZeile := 3, sText := 'offen',  dwFarbe := dwO);
      ELSE                                                             b := VisuHand_Set(stH := pH^, wZeile := 3, sText := '?',      dwFarbe := dwO);
      END_IF
  END_CASE
END_FOR

// Schalter (Toggle) - ausserhalb des Handbetriebs immer zuruecksetzen
IF VISU_HAND.st201.bGesperrt THEN
  VISU_VARS.bgVISUGeblaese[201, cWAND_1] := FALSE;
  VISU_VARS.bgVISUDrosselklappeAUF[201]  := FALSE;
END_IF
IF VISU_HAND.st205.bGesperrt THEN
  VISU_VARS.bgVISUGeblaese[205, cWAND_1] := FALSE;
  VISU_VARS.bgVISUDrosselklappeAUF[205]  := FALSE;
END_IF
IF VISU_HAND.st207.bGesperrt THEN
  VISU_VARS.bgVISUGeblaese[207, cWAND_1] := FALSE;
END_IF

// -------------------------------------------------------------------------------------------
// [101] / [102] SHUTTLE
// -------------------------------------------------------------------------------------------
FOR i := 101 TO 102 DO
  IF i = 101 THEN pH := ADR(VISU_HAND.st101); ELSE pH := ADR(VISU_HAND.st102); END_IF
  pBP := ADR(StationBasisParameter.starrShuttleBasisParameter[i]);
  b := VisuHand_Sperre(stBP := pBP^, stH := pH^, bFaecherwagen := FALSE);
  IF __ISVALIDREF(pBP^.stMKs) THEN
    pH^.abZeileVorhanden[1] := pBP^.stMKs.stStationsAufbau.bGlastransport[cWAND_1];
    pH^.abZeileVorhanden[2] := pBP^.stMKs.stStationsAufbau.bGeblase[cWAND_1];
    pH^.abZeileVorhanden[3] := pBP^.stMKs.stStationsAufbau.bTransportVerstellung[cWAND_1];
    pH^.abZeileVorhanden[4] := pBP^.stMKs.stStationsAufbau.bKippen[cWAND_1];
    pH^.abZeileVorhanden[5] := pBP^.stMKs.stStationsAufbau.bQuerfahrt;
    pH^.abZeileVorhanden[6] := pBP^.stMKs.stStationsAufbau.bDLSSchmiersystem;
    // 7 - 10 Greifer (Ausbaustufe je Wand, in der Visu nur bei 102)
    pH^.abZeileVorhanden[7]  := pBP^.stMKs.stStationsAufbau.bGreifer[cWAND_1];
    pH^.abZeileVorhanden[8]  := pBP^.stMKs.stStationsAufbau.bGreifer[cWAND_1];
    pH^.abZeileVorhanden[9]  := pBP^.stMKs.stStationsAufbau.bGreifer[cWAND_1];
    pH^.abZeileVorhanden[10] := pBP^.stMKs.stStationsAufbau.bGreifer[cWAND_1];
  END_IF
  IF pH^.bGesperrt THEN
    VISU_VARS.bgVISUGeblaese[i, cWAND_1] := FALSE;
  END_IF
  // 1 Riemen
  b := VisuHand_Set(stH := pH^, wZeile := 1,
                     sText   := SEL(abgStationsstatusVisu[i].bSensorEinlauf[1] OR abgStationsstatusVisu[i].bSensorAuslauf[1] OR abgStationsstatusVisu[i].bSensorAuslaufStopp[1], 'frei', 'Glas'),
                     dwFarbe := SEL(abgStationsstatusVisu[i].bSensorEinlauf[1] OR abgStationsstatusVisu[i].bSensorAuslauf[1] OR abgStationsstatusVisu[i].bSensorAuslaufStopp[1], dwGR, dwB));
  // 2 Geblaese
  b := VisuHand_Set(stH := pH^, wZeile := 2, sText := SEL(abgStationsstatusVisu[i].bGeblaeseLaeuft[1], 'aus', 'EIN'), dwFarbe := SEL(abgStationsstatusVisu[i].bGeblaeseLaeuft[1], dwGR, dwB));
  // 3 Oeffnung (Transportverstellung)
  CASE abgStationsstatusVisu[i].epWandverstellungStatus[1] OF
    PneumatikZylinderStatus_EN.eZylinderStellung16mm: b := VisuHand_Set(stH := pH^, wZeile := 3, sText := '16 mm', dwFarbe := dwG);
    PneumatikZylinderStatus_EN.eZylinderStellung23mm: b := VisuHand_Set(stH := pH^, wZeile := 3, sText := '23 mm', dwFarbe := dwG);
    PneumatikZylinderStatus_EN.eZylinderStellung29mm: b := VisuHand_Set(stH := pH^, wZeile := 3, sText := '29 mm', dwFarbe := dwG);
    ELSE                                                b := VisuHand_Set(stH := pH^, wZeile := 3, sText := '?',     dwFarbe := dwO);
  END_CASE
  // 4 Kippen
  CASE abgStationsstatusVisu[i].epKippStatus OF
    Kippen_EN.eKippen_Position_0Grad:    sKipp := '0°';     dwKipp := dwG;
    Kippen_EN.eKippen_Position_84Grad:   sKipp := '84°';    dwKipp := dwG;
    Kippen_EN.eKippen_Position_88_5Grad: sKipp := '88,5°';  dwKipp := dwG;
    Kippen_EN.eKippen_Position_90Grad:   sKipp := '90°';    dwKipp := dwG;
    Kippen_EN.eKippen_Position_96Grad:   sKipp := '96°';    dwKipp := dwG;
    Kippen_EN.eKippen_Fehler:            sKipp := 'Fehler'; dwKipp := dwR;
    ELSE                                   sKipp := 'Zwischen'; dwKipp := dwO;
  END_CASE
  IF abgStationsstatusVisu[i].bKippenFehler THEN dwKipp := dwR; END_IF
  b := VisuHand_Set(stH := pH^, wZeile := 4, sText := sKipp, dwFarbe := dwKipp);
  // 5 Querfahrt
  b := VisuHand_Set(stH := pH^, wZeile := 5,
                     sText   := VisuUeb_MmText(sPrefix := '', rWert := abgStationsstatusVisu[i].rQuerfahrtIstPos, sEinheit := ' mm'),
                     dwFarbe := SEL(abgStationsstatusVisu[i].bQuerfahrtFehler, SEL(abgStationsstatusVisu[i].bQuerfahrtAntriebReferenziert, dwO, dwG), dwR));
  // 6 Schmierung
  b := VisuHand_Set(stH := pH^, wZeile := 6, sText := '', dwFarbe := dwGR);

  // 7 - 10 Greifer (Wand 1)
  IF pH^.abZeileVorhanden[7] THEN
    pGr := ADR(Globale_Bausteine.aShuttle[i].Greifer[cWAND_1]);
    // 7 Greiferachse
    b := VisuHand_Set(stH := pH^, wZeile := 7,
                       sText   := VisuUeb_MmText(sPrefix := '', rWert := pGr^.rpIstPosition, sEinheit := ' mm'),
                       dwFarbe := SEL(pGr^.bpFehler, SEL(pGr^.bpIstInReferenz, dwO, dwG), dwR));
    // 8 Greifer aus- / eingefahren
    IF pGr^.in_bGreiferAusgefahren AND NOT pGr^.in_bGreiferEingefahren THEN
      b := VisuHand_Set(stH := pH^, wZeile := 8, sText := 'ausgefahren', dwFarbe := dwB);
    ELSIF pGr^.in_bGreiferEingefahren AND NOT pGr^.in_bGreiferAusgefahren THEN
      b := VisuHand_Set(stH := pH^, wZeile := 8, sText := 'eingefahren', dwFarbe := dwG);
    ELSE
      b := VisuHand_Set(stH := pH^, wZeile := 8, sText := '?',           dwFarbe := dwO);
    END_IF
    // 9 Greiferzange Auslaufseite (Zange[2] = cZANGE_AUSLAUF im Greifer-Baustein);
    //   nur die Abfrage "offen" wird verwendet (Abfrage "geschlossen" laut MK nicht ausgewertet)
    b := VisuHand_Set(stH := pH^, wZeile := 9,
                       sText   := SEL(pGr^.Zange[2].in_bStatusZylinder_1_Ausgefahren, 'zu', 'offen'),
                       dwFarbe := SEL(pGr^.Zange[2].in_bStatusZylinder_1_Ausgefahren, dwG, dwB));
    // 10 Glasrueckhalter
    b := VisuHand_Set(stH := pH^, wZeile := 10,
                       sText   := SEL(pGr^.bpGlasRueckhalterEingefahren, 'ausgefahren', 'eingefahren'),
                       dwFarbe := SEL(pGr^.bpGlasRueckhalterEingefahren, dwB, dwG));
  END_IF
END_FOR

// -------------------------------------------------------------------------------------------
// [151] / [152] TRANSFERSHUTTLE
// -------------------------------------------------------------------------------------------
FOR i := 151 TO 152 DO
  IF i = 151 THEN pH := ADR(VISU_HAND.st151); ELSE pH := ADR(VISU_HAND.st152); END_IF
  pBP := ADR(StationBasisParameter.starrTransfershuttleBasisParameter[i]);
  b := VisuHand_Sperre(stBP := pBP^, stH := pH^, bFaecherwagen := FALSE);
  IF __ISVALIDREF(pBP^.stMKs) THEN
    pH^.abZeileVorhanden[1] := pBP^.stMKs.stStationsAufbau.bGlastransport[cWAND_1];
    pH^.abZeileVorhanden[2] := pBP^.stMKs.stStationsAufbau.bGlastransport[cWAND_1];
    pH^.abZeileVorhanden[3] := pBP^.stMKs.stStationsAufbau.bDruckluft;
    pH^.abZeileVorhanden[4] := pBP^.stMKs.stStationsAufbau.bDruckluft;
    pH^.abZeileVorhanden[5] := pBP^.stMKs.stStationsAufbau.bQuerfahrt;
    pH^.abZeileVorhanden[6] := pBP^.stMKs.stStationsAufbau.bDLSSchmiersystem;
  END_IF
  IF pH^.bGesperrt THEN
    VISU_VARS.bgVisuTFSRiemenAnheben[i]     := FALSE;
    VISU_VARS.bgVisuTFSAbfrageEinlaufAuf[i] := FALSE;
    VISU_VARS.bgVisuTFSAbfrageEinlaufEin[i] := FALSE;
    VISU_VARS.bgVisuTFSAbfrageAuslaufAuf[i] := FALSE;
    VISU_VARS.bgVisuTFSAbfrageAuslaufEin[i] := FALSE;
  END_IF
  // 1 Riemen
  b := VisuHand_Set(stH := pH^, wZeile := 1,
                     sText   := SEL(abgStationsstatusVisu[i].bSensorEinlauf[1] OR abgStationsstatusVisu[i].bSensorAuslauf[1], 'frei', 'Glas'),
                     dwFarbe := SEL(abgStationsstatusVisu[i].bSensorEinlauf[1] OR abgStationsstatusVisu[i].bSensorAuslauf[1], dwGR, dwB));
  // 2 Riemen Hub (Glastransport angehoben / abgesenkt)
  IF Globale_Bausteine.aTransfershuttles[i].in_bSensorShuttleOben AND NOT Globale_Bausteine.aTransfershuttles[i].in_bSensorShuttleUnten THEN
    b := VisuHand_Set(stH := pH^, wZeile := 2, sText := 'angehoben', dwFarbe := dwB);
  ELSIF Globale_Bausteine.aTransfershuttles[i].in_bSensorShuttleUnten AND NOT Globale_Bausteine.aTransfershuttles[i].in_bSensorShuttleOben THEN
    b := VisuHand_Set(stH := pH^, wZeile := 2, sText := 'abgesenkt', dwFarbe := dwG);
  ELSE
    b := VisuHand_Set(stH := pH^, wZeile := 2, sText := '?', dwFarbe := dwO);
  END_IF
  // 3 / 4 Scheibenabfrage Einlauf / Auslauf
  b := VisuHand_Set(stH := pH^, wZeile := 3, sText := SEL(abgStationsstatusVisu[i].bSensorEinlauf[1], 'frei', 'belegt'), dwFarbe := SEL(abgStationsstatusVisu[i].bSensorEinlauf[1], dwGR, dwB));
  b := VisuHand_Set(stH := pH^, wZeile := 4, sText := SEL(abgStationsstatusVisu[i].bSensorAuslauf[1], 'frei', 'belegt'), dwFarbe := SEL(abgStationsstatusVisu[i].bSensorAuslauf[1], dwGR, dwB));
  // 5 Querfahrt
  b := VisuHand_Set(stH := pH^, wZeile := 5,
                     sText   := VisuUeb_MmText(sPrefix := '', rWert := abgStationsstatusVisu[i].rQuerfahrtIstPos, sEinheit := ' mm'),
                     dwFarbe := SEL(abgStationsstatusVisu[i].bQuerfahrtFehler, SEL(abgStationsstatusVisu[i].bQuerfahrtAntriebReferenziert, dwO, dwG), dwR));
  // 6 Schmierung
  b := VisuHand_Set(stH := pH^, wZeile := 6, sText := '', dwFarbe := dwGR);
END_FOR

// -------------------------------------------------------------------------------------------
// [301] - [305] FAECHERWAGEN (Variante Einfach: Rolltor, Arretierung = Gegenhalter)
// -------------------------------------------------------------------------------------------
FOR i := 301 TO 305 DO
  pBP := ADR(StationBasisParameter.starrFaecherwagenBasisParameter[i]);
  b := VisuHand_Sperre(stBP := pBP^, stH := VISU_HAND.astFW[i], bFaecherwagen := TRUE);
  IF __ISVALIDREF(pBP^.stMKs) THEN
    VISU_HAND.astFW[i].abZeileVorhanden[1] := pBP^.stMKs.stStationsAufbau.bRolltor;
    VISU_HAND.astFW[i].abZeileVorhanden[2] := TRUE;
  END_IF

  // Rolltor-Schalter gegenseitig ausschliessen, ausserhalb des Handbetriebs zuruecksetzen
  artlRolltorHoch[i](CLK := VISU_VARS.bgVISUFWRolltorHoch[i]);
  artlRolltorRunter[i](CLK := VISU_VARS.bgVISUFWRolltorRunter[i]);
  IF artlRolltorHoch[i].Q THEN   VISU_VARS.bgVISUFWRolltorRunter[i] := FALSE; END_IF
  IF artlRolltorRunter[i].Q THEN VISU_VARS.bgVISUFWRolltorHoch[i]   := FALSE; END_IF
  IF VISU_HAND.astFW[i].bGesperrt THEN
    VISU_VARS.bgVISUFWRolltorHoch[i]   := FALSE;
    VISU_VARS.bgVISUFWRolltorRunter[i] := FALSE;
  END_IF

  // 1 Rolltor
  IF VISU_VARS.astgFaecherwagenstatusVisu[i].bRolltorOben THEN
    b := VisuHand_Set(stH := VISU_HAND.astFW[i], wZeile := 1, sText := 'oben',  dwFarbe := dwG);
  ELSIF VISU_VARS.astgFaecherwagenstatusVisu[i].bRolltorUnten THEN
    b := VisuHand_Set(stH := VISU_HAND.astFW[i], wZeile := 1, sText := 'unten', dwFarbe := dwG);
  ELSE
    b := VisuHand_Set(stH := VISU_HAND.astFW[i], wZeile := 1, sText := '?',     dwFarbe := dwO);
  END_IF
  // 2 Gegenhalter (Arretierung): Endlage 1 = offen, 2 = geschlossen
  IF VISU_VARS.astgFaecherwagenstatusVisu[i].abEndlage[1] THEN
    b := VisuHand_Set(stH := VISU_HAND.astFW[i], wZeile := 2, sText := 'offen', dwFarbe := dwG);
  ELSIF VISU_VARS.astgFaecherwagenstatusVisu[i].abEndlage[2] THEN
    b := VisuHand_Set(stH := VISU_HAND.astFW[i], wZeile := 2, sText := 'zu',    dwFarbe := dwG);
  ELSE
    b := VisuHand_Set(stH := VISU_HAND.astFW[i], wZeile := 2, sText := '?',     dwFarbe := dwO);
  END_IF
END_FOR
END_PROGRAM

(* ---- VisuUebersicht_PRG.prg.st ---- *)
(* METADATA
{
	"v3Meta": {
		"objectGuid": "ba53d487-b3e7-4729-ab5c-8ab03e7357e2"
	}
}
*)
PROGRAM VisuUebersicht_PRG
VAR
  bBlink        : BOOL;
  bLernen       : BOOL;
  bSK1, bSK2    : BOOL;
  bSK3, bSK4    : BOOL;
  bStoerung     : BOOL;
  wAnzStoerung  : WORD;
  sKipp         : STRING(40);
  sDreh         : STRING(20);
  sTitel        : STRING(40);
  pKarte        : POINTER TO VisuUeb_Station_ST;
  pAchse        : POINTER TO VisuUeb_Achse_ST;
  pInit         : POINTER TO BOOL;
  pMin, pMax    : POINTER TO REAL;
  rQuerMin      : REAL;
  rQuerMax      : REAL;
  bDummy        : BOOL;
  wIdx          : WORD;
  sNr           : STRING(5);
END_VAR
// *************************************************************************************************
// DATENAUFBEREITUNG FUER DIE VISU "Anlagenuebersicht"
// - Visu verwendet ausschliesslich die Variablen aus VISU_UEBERSICHT (Texte, Farben, Pixel)
// *************************************************************************************************
bBlink  := Global_Vars.gbFlashbit05sec;
bLernen := VISU_UEBERSICHT.bSkalierungNeuLernen;
VISU_UEBERSICHT.bSkalierungNeuLernen := FALSE;

// -------------------------------------------------------------------------------------------
// KOPFZEILE
// -------------------------------------------------------------------------------------------
bSK1 := Globale_Bausteine.Sicherheitskreis[1].bpSicherheitskreisGeschlossen;
bSK2 := Globale_Bausteine.Sicherheitskreis[2].bpSicherheitskreisGeschlossen;
bSK3 := Globale_Bausteine.Sicherheitskreis[3].bpSicherheitskreisGeschlossen;
bSK4 := Globale_Bausteine.Sicherheitskreis[4].bpSicherheitskreisGeschlossen;

bDummy := VisuUeb_Lampe(stLampe := VISU_UEBERSICHT.stAutomatik,      sText := SEL(Global_Vars.M_Automatik_Aktiv[1], 'HAND', 'AUTOMATIK'), bOK := Global_Vars.M_Automatik_Aktiv[1], bWarnung := TRUE, bNeutral := FALSE);
bDummy := VisuUeb_Lampe(stLampe := VISU_UEBERSICHT.stSK1,            sText := SEL(bSK1, 'SK 1 offen', 'SK 1 zu'), bOK := bSK1, bWarnung := TRUE, bNeutral := FALSE);
bDummy := VisuUeb_Lampe(stLampe := VISU_UEBERSICHT.stSK2,            sText := SEL(bSK2, 'SK 2 offen', 'SK 2 zu'), bOK := bSK2, bWarnung := TRUE, bNeutral := FALSE);
bDummy := VisuUeb_Lampe(stLampe := VISU_UEBERSICHT.stSK3,            sText := SEL(bSK3, 'SK 3 offen', 'SK 3 zu'), bOK := bSK3, bWarnung := TRUE, bNeutral := FALSE);
bDummy := VisuUeb_Lampe(stLampe := VISU_UEBERSICHT.stSK4,            sText := SEL(bSK4, 'SK 4 offen', 'SK 4 zu'), bOK := bSK4, bWarnung := TRUE, bNeutral := FALSE);
// Tueren: je Tuer eine Anzeige (zu = gruen, Anforderung = orange blinkend, offen = rot)
FOR wIdx := 1 TO VISU_UEBERSICHT.cMAX_TUEREN DO
  VISU_UEBERSICHT.abTuerVorhanden[wIdx] := (wIdx >= Stations_Konfig.cERSTE_TUER) AND (wIdx <= Stations_Konfig.cLETZTE_TUER);
  IF VISU_UEBERSICHT.abTuerVorhanden[wIdx] THEN
    sNr := WORD_TO_STRING(wIdx);
    IF Globale_Bausteine.aTuer[wIdx].bpStatusTuerNichtGeschlossen THEN
      VISU_UEBERSICHT.astTuer[wIdx].sText   := CONCAT(CONCAT('Tür ', sNr), ' offen');
      VISU_UEBERSICHT.astTuer[wIdx].dwFarbe := VISU_UEBERSICHT.cFARBE_ROT;
    ELSIF Globale_Bausteine.aTuer[wIdx].bpAnforderungZumTuerOffnenGestellt THEN
      VISU_UEBERSICHT.astTuer[wIdx].sText   := CONCAT(CONCAT('Tür ', sNr), ' Anford.');
      VISU_UEBERSICHT.astTuer[wIdx].dwFarbe := SEL(bBlink, VISU_UEBERSICHT.cFARBE_GRAU, VISU_UEBERSICHT.cFARBE_ORANGE);
    ELSE
      VISU_UEBERSICHT.astTuer[wIdx].sText   := CONCAT(CONCAT('Tür ', sNr), ' zu');
      VISU_UEBERSICHT.astTuer[wIdx].dwFarbe := VISU_UEBERSICHT.cFARBE_GRUEN;
    END_IF
  END_IF
END_FOR

// Durchgaenge
FOR wIdx := 1 TO VISU_UEBERSICHT.cMAX_DURCHGAENGE DO
  VISU_UEBERSICHT.abDurchgangVorhanden[wIdx] := (wIdx >= Stations_Konfig.cERSTER_DURCHGANG) AND (wIdx <= Stations_Konfig.cLETZTER_DURCHGANG);
  IF VISU_UEBERSICHT.abDurchgangVorhanden[wIdx] THEN
    sNr := WORD_TO_STRING(wIdx);
    IF Globale_Bausteine.aDurchgang[wIdx].bpStatusDurchgangNichtGeschlossen THEN
      VISU_UEBERSICHT.astDurchgang[wIdx].sText   := CONCAT(CONCAT('Durchgang ', sNr), ' offen');
      VISU_UEBERSICHT.astDurchgang[wIdx].dwFarbe := VISU_UEBERSICHT.cFARBE_ROT;
    ELSIF Globale_Bausteine.aDurchgang[wIdx].bpAnforderungZumDurchgangOffnenGestellt THEN
      VISU_UEBERSICHT.astDurchgang[wIdx].sText   := CONCAT(CONCAT('Durchgang ', sNr), ' Anf.');
      VISU_UEBERSICHT.astDurchgang[wIdx].dwFarbe := SEL(bBlink, VISU_UEBERSICHT.cFARBE_GRAU, VISU_UEBERSICHT.cFARBE_ORANGE);
    ELSE
      VISU_UEBERSICHT.astDurchgang[wIdx].sText   := CONCAT(CONCAT('Durchgang ', sNr), ' zu');
      VISU_UEBERSICHT.astDurchgang[wIdx].dwFarbe := VISU_UEBERSICHT.cFARBE_GRUEN;
    END_IF
  END_IF
END_FOR
bDummy := VisuUeb_Lampe(stLampe := VISU_UEBERSICHT.stDruckluft,      sText := 'Druckluft',     bOK := StatusAnlage.abpDruckluftOK[1], bWarnung := FALSE, bNeutral := FALSE);
bDummy := VisuUeb_Lampe(stLampe := VISU_UEBERSICHT.stSchaltschrank,  sText := 'Schaltschrank', bOK := StatusAnlage.bpAnlageOK, bWarnung := FALSE, bNeutral := FALSE);
bDummy := VisuUeb_Lampe(stLampe := VISU_UEBERSICHT.stEtherCAT,       sText := 'EtherCAT',      bOK := Global_Vars.bgEtherCatOK, bWarnung := FALSE, bNeutral := FALSE);
bDummy := VisuUeb_Lampe(stLampe := VISU_UEBERSICHT.stInit,           sText := 'Init',          bOK := Global_Vars.M_Init_Ok, bWarnung := TRUE, bNeutral := FALSE);
bDummy := VisuUeb_Lampe(stLampe := VISU_UEBERSICHT.stMMI,            sText := 'MMI',           bOK := MMI_Vars.bgMMIOK OR Global_Vars.bgMMIBruecken, bWarnung := Global_Vars.bgMMIBruecken, bNeutral := FALSE);
bDummy := VisuUeb_Lampe(stLampe := VISU_UEBERSICHT.stBetriebsstop,   sText := SEL(Globale_Bausteine.Stop_Baustein.abpBetriebsstop[1], 'Betrieb', 'BETRIEBSSTOP'), bOK := NOT Globale_Bausteine.Stop_Baustein.abpBetriebsstop[1], bWarnung := FALSE, bNeutral := FALSE);
bDummy := VisuUeb_Lampe(stLampe := VISU_UEBERSICHT.stInbetriebnahme, sText := 'IBN-Modus',     bOK := FALSE, bWarnung := TRUE, bNeutral := NOT Global_Vars.bgInbetriebnahmeBit);

// -------------------------------------------------------------------------------------------
// STATIONEN
// -------------------------------------------------------------------------------------------
wAnzStoerung := 0;

// [501] Einlauf Fremdanlage (VSG)
IF VisuUeb_Station(stBP := StationBasisParameter.starrFremdanlageEinlaufStationBasisParameter[501], stKarte := VISU_UEBERSICHT.st501, sTitel := '501  Einlauf VSG', bBlink := bBlink, bReferenzRelevant := FALSE, bGlasZusatz := FALSE) THEN wAnzStoerung := wAnzStoerung + 1; END_IF
VISU_UEBERSICHT.st501.sInfo1 := SEL(VISU_VARS.abgVISUFreigabeFremdanlage[501], 'Freigabe Visu: aus', 'Freigabe Visu: EIN');
VISU_UEBERSICHT.st501.sInfo2 := '';
VISU_UEBERSICHT.st501.sInfo3 := '';

// [201] - [208] Stationen der Zufuehrung: Karte, Glas und Sensoren
FOR wIdx := 201 TO 208 DO
  CASE wIdx OF
    201: pKarte := ADR(VISU_UEBERSICHT.st201); sTitel := '201  Anlegetisch';
    202: pKarte := ADR(VISU_UEBERSICHT.st202); sTitel := '202  Förderer';
    203: pKarte := ADR(VISU_UEBERSICHT.st203); sTitel := '203  Förderer';
    204: pKarte := ADR(VISU_UEBERSICHT.st204); sTitel := '204  Eckübergabe';
    205: pKarte := ADR(VISU_UEBERSICHT.st205); sTitel := '205  Anlegetisch';
    206: pKarte := ADR(VISU_UEBERSICHT.st206); sTitel := '206  Kipptisch';
    207: pKarte := ADR(VISU_UEBERSICHT.st207); sTitel := '207  Drehstation';
    208: pKarte := ADR(VISU_UEBERSICHT.st208); sTitel := '208  Anlegewand';
  END_CASE
  IF VisuUeb_Station(stBP := StationBasisParameter.starrStationBasisParameter[wIdx], stKarte := pKarte^, sTitel := sTitel, bBlink := bBlink, bReferenzRelevant := TRUE,
                      bGlasZusatz := abgStationsstatusVisu[wIdx].bSensorEinlauf[1] OR abgStationsstatusVisu[wIdx].bSensorAuslauf[1]) THEN wAnzStoerung := wAnzStoerung + 1; END_IF
  pKarte^.dwSensorEinlauf      := VisuUeb_Sensor(abgStationsstatusVisu[wIdx].bSensorEinlauf[1]);
  pKarte^.dwSensorEinlaufVorab := VisuUeb_Sensor(abgStationsstatusVisu[wIdx].bSensorEinlaufVorab[1]);
  pKarte^.dwSensorAuslaufVorab := VisuUeb_Sensor(abgStationsstatusVisu[wIdx].bSensorAuslaufVorab[1]);
  pKarte^.dwSensorAuslauf      := VisuUeb_Sensor(abgStationsstatusVisu[wIdx].bSensorAuslauf[1]);
  pKarte^.sInfo1 := '';  pKarte^.dwInfo1Farbe := VISU_UEBERSICHT.cFARBE_TEXT;
  pKarte^.sInfo2 := '';  pKarte^.dwInfo2Farbe := VISU_UEBERSICHT.cFARBE_TEXT;
  pKarte^.sInfo3 := '';  pKarte^.dwInfo3Farbe := VISU_UEBERSICHT.cFARBE_TEXT;

  // Anlegetisch: Messachse, Anschlag, Hubrahmen, Ampel
  IF wIdx = 201 OR wIdx = 205 THEN
    pKarte^.sInfo1 := VisuUeb_MmText(sPrefix := 'Messachse ', rWert := abgStationsstatusVisu[wIdx].rMessachseIstPos);
    pKarte^.dwInfo1Farbe := SEL(abgStationsstatusVisu[wIdx].bMessachseFehler, VISU_UEBERSICHT.cFARBE_TEXT, VISU_UEBERSICHT.cFARBE_ROT);
    pKarte^.sInfo2 := CONCAT(CONCAT('Anschlag ', SEL(abgStationsstatusVisu[wIdx].bAnschlagSensorAusgefahren, SEL(abgStationsstatusVisu[wIdx].bAnschlagSensorEingefahren, '?', 'unten'), 'oben')),
                             CONCAT(' | Hubrahmen ', SEL(abgStationsstatusVisu[wIdx].bHubpaletteSensorAusgefahren, SEL(abgStationsstatusVisu[wIdx].bHubpaletteSensorEingefahren, '?', 'unten'), 'oben')));
    pKarte^.dwInfo2Farbe := SEL(abgStationsstatusVisu[wIdx].bAnschlagFehler OR abgStationsstatusVisu[wIdx].bHubpaletteFehler, VISU_UEBERSICHT.cFARBE_TEXT, VISU_UEBERSICHT.cFARBE_ROT);
    pKarte^.sInfo3 := CONCAT('Ampel ', SEL(abgStationsstatusVisu[wIdx].bAmpelRot, SEL(abgStationsstatusVisu[wIdx].bAmpelGruen, 'aus', 'grün'), 'rot'));
  END_IF
END_FOR

// [206] Kipptisch
CASE abgStationsstatusVisu[206].epKippStatus OF
  Kippen_EN.eKippen_Position_0Grad:    sKipp := '0°';
  Kippen_EN.eKippen_Position_84Grad:   sKipp := '84°';
  Kippen_EN.eKippen_Position_88_5Grad: sKipp := '88,5°';
  Kippen_EN.eKippen_Position_90Grad:   sKipp := '90°';
  Kippen_EN.eKippen_Position_96Grad:   sKipp := '96°';
  Kippen_EN.eKippen_Fehler:            sKipp := 'FEHLER';
  ELSE                                   sKipp := 'Zwischenpos.';
END_CASE
VISU_UEBERSICHT.st206.sInfo1 := CONCAT(CONCAT('Kippen ', sKipp), VisuUeb_MmText(sPrefix := '  (', rWert := abgStationsstatusVisu[206].rKippenIstPos, sEinheit := ')'));
VISU_UEBERSICHT.st206.dwInfo1Farbe := SEL(abgStationsstatusVisu[206].bKippenFehler OR NOT abgStationsstatusVisu[206].bKippenAntriebReferenziert, VISU_UEBERSICHT.cFARBE_TEXT, VISU_UEBERSICHT.cFARBE_ROT);
VISU_UEBERSICHT.st206.sInfo2 := SEL(abgStationsstatusVisu[206].bKippenMinEndschalter OR abgStationsstatusVisu[206].bKippenMaxEndschalter, 'Endschalter frei', 'ENDSCHALTER BELEGT');
VISU_UEBERSICHT.st206.dwInfo2Farbe := SEL(abgStationsstatusVisu[206].bKippenMinEndschalter OR abgStationsstatusVisu[206].bKippenMaxEndschalter, VISU_UEBERSICHT.cFARBE_TEXT, VISU_UEBERSICHT.cFARBE_ROT);

// [207] Drehstation
CASE abgStationsstatusVisu[207].epDrehIstPosition OF
  Drehen_EN.eDrehPosition0Grad:   sDreh := '0°';
  Drehen_EN.eDrehPosition90Grad:  sDreh := '90°';
  Drehen_EN.eDrehPosition180Grad: sDreh := '180°';
  Drehen_EN.eDrehPosition270Grad: sDreh := '270°';
  ELSE                              sDreh := 'Zwischenpos.';
END_CASE
VISU_UEBERSICHT.st207.sInfo1 := CONCAT(CONCAT('Drehen ', sDreh), VisuUeb_MmText(sPrefix := '  (', rWert := abgStationsstatusVisu[207].rDrehenIstPos, sEinheit := ')'));
VISU_UEBERSICHT.st207.dwInfo1Farbe := SEL(abgStationsstatusVisu[207].bDrehenFehler OR NOT abgStationsstatusVisu[207].bDrehenAntriebReferenziert, VISU_UEBERSICHT.cFARBE_TEXT, VISU_UEBERSICHT.cFARBE_ROT);
VISU_UEBERSICHT.st207.sInfo2 := CONCAT('Arretierung ', SEL(abgStationsstatusVisu[207].bDrehenArretierungAusgefahren, SEL(abgStationsstatusVisu[207].bDrehenArretierungEingefahren, '?', 'eingefahren'), 'ausgefahren'));
VISU_UEBERSICHT.st207.sInfo3 := SEL(EV_ToPLC_b207_geschlossen, 'Durchfassperre 208 OFFEN', 'Durchfassperre 208 zu');
VISU_UEBERSICHT.st207.dwInfo3Farbe := SEL(EV_ToPLC_b207_geschlossen, VISU_UEBERSICHT.cFARBE_ROT, VISU_UEBERSICHT.cFARBE_TEXT);

// [208] Anlegewand
VISU_UEBERSICHT.st208.sInfo1 := VisuUeb_MmText(sPrefix := 'Messachse ', rWert := abgStationsstatusVisu[208].rMessachseIstPos);
VISU_UEBERSICHT.st208.dwInfo1Farbe := SEL(abgStationsstatusVisu[208].bMessachseFehler, VISU_UEBERSICHT.cFARBE_TEXT, VISU_UEBERSICHT.cFARBE_ROT);
VISU_UEBERSICHT.st208.sInfo2 := CONCAT('Ampel ', SEL(abgStationsstatusVisu[208].bAmpelRot, SEL(abgStationsstatusVisu[208].bAmpelGruen, 'aus', 'grün'), 'rot'));

// [101] / [102] Shuttle
// Beide Querfahrten gehoeren zum selben Koordinatensystem: gemeinsamer Darstellungsbereich,
// damit gleiche Position = gleiche Hoehe in der Visu (Bereich der Vorrunde)
IF VISU_UEBERSICHT.bSkalierung101Init AND VISU_UEBERSICHT.bSkalierung102Init THEN
  rQuerMin := MIN(VISU_UEBERSICHT.rMin101, VISU_UEBERSICHT.rMin102);
  rQuerMax := MAX(VISU_UEBERSICHT.rMax101, VISU_UEBERSICHT.rMax102);
ELSE
  rQuerMin := 0.0;
  rQuerMax := 0.0;
END_IF
FOR wIdx := 101 TO 102 DO
  IF wIdx = 101 THEN
    pKarte := ADR(VISU_UEBERSICHT.st101); pAchse := ADR(VISU_UEBERSICHT.stAchse101); sTitel := '101  Shuttle';
    pInit := ADR(VISU_UEBERSICHT.bSkalierung101Init); pMin := ADR(VISU_UEBERSICHT.rMin101); pMax := ADR(VISU_UEBERSICHT.rMax101);
  ELSE
    pKarte := ADR(VISU_UEBERSICHT.st102); pAchse := ADR(VISU_UEBERSICHT.stAchse102); sTitel := '102  Shuttle';
    pInit := ADR(VISU_UEBERSICHT.bSkalierung102Init); pMin := ADR(VISU_UEBERSICHT.rMin102); pMax := ADR(VISU_UEBERSICHT.rMax102);
  END_IF
  IF VisuUeb_Station(stBP := StationBasisParameter.starrShuttleBasisParameter[wIdx], stKarte := pKarte^, sTitel := sTitel, bBlink := bBlink, bReferenzRelevant := TRUE,
                      bGlasZusatz := abgStationsstatusVisu[wIdx].bSensorEinlauf[1] OR abgStationsstatusVisu[wIdx].bSensorAuslauf[1] OR abgStationsstatusVisu[wIdx].bSensorAuslaufStopp[1]) THEN wAnzStoerung := wAnzStoerung + 1; END_IF
  pKarte^.dwSensorEinlauf      := VisuUeb_Sensor(abgStationsstatusVisu[wIdx].bSensorEinlauf[1]);
  pKarte^.dwSensorEinlaufVorab := VisuUeb_Sensor(abgStationsstatusVisu[wIdx].bSensorEinlaufVorab[1]);
  pKarte^.dwSensorAuslaufVorab := VisuUeb_Sensor(abgStationsstatusVisu[wIdx].bSensorAuslaufVorab[1]);
  pKarte^.dwSensorAuslauf      := VisuUeb_Sensor(abgStationsstatusVisu[wIdx].bSensorAuslauf[1]);
  pKarte^.dwSensorAuslaufStopp := VisuUeb_Sensor(abgStationsstatusVisu[wIdx].bSensorAuslaufStopp[1]);
  CASE abgStationsstatusVisu[wIdx].epKippStatus OF
    Kippen_EN.eKippen_Position_0Grad:    sKipp := 'Kippen 0°';
    Kippen_EN.eKippen_Position_84Grad:   sKipp := 'Kippen 84°';
    Kippen_EN.eKippen_Position_88_5Grad: sKipp := 'Kippen 88,5°';
    Kippen_EN.eKippen_Position_90Grad:   sKipp := 'Kippen 90°';
    Kippen_EN.eKippen_Position_96Grad:   sKipp := 'Kippen 96°';
    Kippen_EN.eKippen_Fehler:            sKipp := 'Kippen FEHLER';
    ELSE                                   sKipp := 'Kippen Zwischenpos.';
  END_CASE
  IF ( Globale_Bausteine.aShuttle[wIdx].Kippen.bpAktivieren ) THEN
    pKarte^.sInfo1 := CONCAT(sKipp, SEL(abgStationsstatusVisu[wIdx].bGeblaeseLaeuft[1], ' | Gebläse aus', ' | Gebläse EIN'));
  ELSE
    pKarte^.sInfo1 := SEL(abgStationsstatusVisu[wIdx].bGeblaeseLaeuft[1], 'Gebläse aus', 'Gebläse EIN');
  END_IF
  pKarte^.dwInfo1Farbe := SEL(abgStationsstatusVisu[wIdx].bKippenFehler AND Globale_Bausteine.aShuttle[wIdx].Kippen.bpAktivieren, VISU_UEBERSICHT.cFARBE_TEXT, VISU_UEBERSICHT.cFARBE_ROT);

  // Fahrwegsgrenzen aus dem Antrieb (Software-Endlagen)
  IF __ISVALIDREF(Globale_Bausteine.aShuttle[wIdx].Querfahrt.Antrieb) THEN
    pMin^  := Globale_Bausteine.aShuttle[wIdx].Querfahrt.Antrieb.rpMinPosition;
    pMax^  := Globale_Bausteine.aShuttle[wIdx].Querfahrt.Antrieb.rpMaxPosition;
    pInit^ := TRUE;
  END_IF
  VisuUeb_Achse(stAchse := pAchse^, bInit := pInit^, rMin := pMin^, rMax := pMax^,
                 rIst            := abgStationsstatusVisu[wIdx].rQuerfahrtIstPos,
                 rZiel           := Globale_Bausteine.aShuttle[wIdx].Querfahrt.rpDestinationPosition,
                 rSpeed          := Globale_Bausteine.aShuttle[wIdx].Querfahrt.rpAktSpeed,
                 bPositionierung := Globale_Bausteine.aShuttle[wIdx].Querfahrt.bpPositionierungAktiv,
                 bReferenziert   := abgStationsstatusVisu[wIdx].bQuerfahrtAntriebReferenziert,
                 bFehler         := abgStationsstatusVisu[wIdx].bQuerfahrtFehler,
                 bMinEnd         := abgStationsstatusVisu[wIdx].bQuerfahrtMinEndschalter,
                 bMaxEnd         := abgStationsstatusVisu[wIdx].bQuerfahrtMaxEndschalter,
                 bNeuLernen      := bLernen,
                 bBlink          := bBlink,
                 rSkalaMin       := rQuerMin,
                 rSkalaMax       := rQuerMax);
  pKarte^.sInfo2 := pAchse^.sIstPos;
  pKarte^.sInfo3 := pAchse^.sZielPos;
END_FOR

// [151] / [152] Transfershuttle
FOR wIdx := 151 TO 152 DO
  IF wIdx = 151 THEN
    pKarte := ADR(VISU_UEBERSICHT.st151); pAchse := ADR(VISU_UEBERSICHT.stAchse151); sTitel := '151  Transfershuttle';
    pInit := ADR(VISU_UEBERSICHT.bSkalierung151Init); pMin := ADR(VISU_UEBERSICHT.rMin151); pMax := ADR(VISU_UEBERSICHT.rMax151);
  ELSE
    pKarte := ADR(VISU_UEBERSICHT.st152); pAchse := ADR(VISU_UEBERSICHT.stAchse152); sTitel := '152  Transfershuttle';
    pInit := ADR(VISU_UEBERSICHT.bSkalierung152Init); pMin := ADR(VISU_UEBERSICHT.rMin152); pMax := ADR(VISU_UEBERSICHT.rMax152);
  END_IF
  IF VisuUeb_Station(stBP := StationBasisParameter.starrTransfershuttleBasisParameter[wIdx], stKarte := pKarte^, sTitel := sTitel, bBlink := bBlink, bReferenzRelevant := TRUE,
                      bGlasZusatz := abgStationsstatusVisu[wIdx].bSensorEinlauf[1] OR abgStationsstatusVisu[wIdx].bSensorAuslauf[1]) THEN wAnzStoerung := wAnzStoerung + 1; END_IF
  pKarte^.dwSensorEinlauf      := VisuUeb_Sensor(abgStationsstatusVisu[wIdx].bSensorEinlauf[1]);
  pKarte^.dwSensorEinlaufVorab := VisuUeb_Sensor(FALSE, FALSE);
  pKarte^.dwSensorAuslaufVorab := VisuUeb_Sensor(FALSE, FALSE);
  pKarte^.dwSensorAuslauf      := VisuUeb_Sensor(abgStationsstatusVisu[wIdx].bSensorAuslauf[1]);
  pKarte^.sInfo1 := SEL(Global_Vars.abgVerfahrfreigabeShuttle[wIdx], 'Verfahrfreigabe: NEIN', 'Verfahrfreigabe: ja');
  pKarte^.dwInfo1Farbe := SEL(Global_Vars.abgVerfahrfreigabeShuttle[wIdx], VISU_UEBERSICHT.cFARBE_ORANGE, VISU_UEBERSICHT.cFARBE_TEXT);

  // Fahrwegsgrenzen aus dem Antrieb (Software-Endlagen)
  IF __ISVALIDREF(Globale_Bausteine.aTransfershuttles[wIdx].Querfahrt.Antrieb) THEN
    pMin^  := Globale_Bausteine.aTransfershuttles[wIdx].Querfahrt.Antrieb.rpMinPosition;
    pMax^  := Globale_Bausteine.aTransfershuttles[wIdx].Querfahrt.Antrieb.rpMaxPosition;
    pInit^ := TRUE;
  END_IF
  VisuUeb_Achse(stAchse := pAchse^, bInit := pInit^, rMin := pMin^, rMax := pMax^,
                 rIst            := abgStationsstatusVisu[wIdx].rQuerfahrtIstPos,
                 rZiel           := Globale_Bausteine.aTransfershuttles[wIdx].Querfahrt.rpDestinationPosition,
                 rSpeed          := Globale_Bausteine.aTransfershuttles[wIdx].Querfahrt.rpAktSpeed,
                 bPositionierung := Globale_Bausteine.aTransfershuttles[wIdx].Querfahrt.bpPositionierungAktiv,
                 bReferenziert   := abgStationsstatusVisu[wIdx].bQuerfahrtAntriebReferenziert,
                 bFehler         := abgStationsstatusVisu[wIdx].bQuerfahrtFehler,
                 bMinEnd         := abgStationsstatusVisu[wIdx].bQuerfahrtMinEndschalter,
                 bMaxEnd         := abgStationsstatusVisu[wIdx].bQuerfahrtMaxEndschalter,
                 bNeuLernen      := bLernen,
                 bBlink          := bBlink,
                 rSkalaMin       := 0.0,
                 rSkalaMax       := 0.0);
  pKarte^.sInfo2 := pAchse^.sIstPos;
  pKarte^.sInfo3 := CONCAT(CONCAT(pAchse^.sZielPos, '   '), pAchse^.sSpeed);
END_FOR

// [301] - [305] Faecherwagen
FOR wIdx := 301 TO 305 DO
  CASE wIdx OF
    301: pKarte := ADR(VISU_UEBERSICHT.st301);
    302: pKarte := ADR(VISU_UEBERSICHT.st302);
    303: pKarte := ADR(VISU_UEBERSICHT.st303);
    304: pKarte := ADR(VISU_UEBERSICHT.st304);
    305: pKarte := ADR(VISU_UEBERSICHT.st305);
  END_CASE
  sTitel := CONCAT(WORD_TO_STRING(wIdx), '  Fächerwagen');
  IF VisuUeb_Station(stBP := StationBasisParameter.starrFaecherwagenBasisParameter[wIdx], stKarte := pKarte^, sTitel := sTitel, bBlink := bBlink, bReferenzRelevant := FALSE,
                      bGlasZusatz := VISU_VARS.astgFaecherwagenstatusVisu[wIdx].bStatusStationInBeladePosition) THEN wAnzStoerung := wAnzStoerung + 1; END_IF
  pKarte^.sInfo1 := CONCAT(SEL(VISU_VARS.astgFaecherwagenstatusVisu[wIdx].bWagenErkannt, 'Kein Fächerwagen', 'Fächerwagen vorhanden'),
                           SEL(VISU_VARS.astgFaecherwagenstatusVisu[wIdx].bRolltorUnten, SEL(VISU_VARS.astgFaecherwagenstatusVisu[wIdx].bRolltorOben, ' | Rolltor ?', ' | Rolltor oben'), ' | Rolltor unten'));
  pKarte^.dwInfo1Farbe := VISU_UEBERSICHT.cFARBE_TEXT;
  IF VISU_VARS.astgFaecherwagenstatusVisu[wIdx].bAuftragAktiv THEN
    pKarte^.sInfo2 := 'Ein-/Ausschleusen aktiv';
    pKarte^.dwInfo2Farbe := VISU_UEBERSICHT.cFARBE_BLAU;
  ELSE
    pKarte^.sInfo2 := SEL(VISU_VARS.astgFaecherwagenstatusVisu[wIdx].bStatusStationInBeladePosition, 'Wagen nicht in Beladeposition', 'Wagen in Beladeposition');
    pKarte^.dwInfo2Farbe := SEL(VISU_VARS.astgFaecherwagenstatusVisu[wIdx].bStatusStationInBeladePosition, VISU_UEBERSICHT.cFARBE_TEXT, VISU_UEBERSICHT.cFARBE_GRUEN);
  END_IF
END_FOR

// -------------------------------------------------------------------------------------------
// SAMMELMELDUNG
// -------------------------------------------------------------------------------------------
bStoerung := wAnzStoerung > 0;
IF bStoerung THEN
  VISU_UEBERSICHT.sStoerungen       := CONCAT(WORD_TO_STRING(wAnzStoerung), SEL(wAnzStoerung = 1, ' Stationen in Störung', ' Station in Störung'));
  VISU_UEBERSICHT.dwStoerungenFarbe := SEL(bBlink, 16#FFA83232, VISU_UEBERSICHT.cFARBE_ROT);
ELSE
  VISU_UEBERSICHT.sStoerungen       := 'Keine Störung';
  VISU_UEBERSICHT.dwStoerungenFarbe := VISU_UEBERSICHT.cFARBE_GRUEN;
END_IF
END_PROGRAM
